Fanuc KAREL source: kd00021.KL

-- PROVISIONAL review KL for V770-1; original PC SHA256 95456d19cd32df8edbdbc64815a97ad4388cbccc3273ca6e1f46dacfe11a0894
-- Incomplete behavior may be omitted. Consult companion uncertainty JSON. Do not deploy.
PROGRAM KD00021
%NOLOCKGROUP
BEGIN
  -- UNRESOLVED_PC offsets 5-17; opcodes 21,23
  -- UNRESOLVED_PC offsets 22-26; opcodes 7F
END KD00021
